# EPICS autosave request: iocs/motor/xps-ioc/db/XPSPositionCompare_settings.req
$(P)$(R)PositionCompareMode
$(P)$(R)PositionCompareMinPosition
$(P)$(R)PositionCompareMaxPosition
$(P)$(R)PositionCompareStepSize
$(P)$(R)PositionComparePulseWidth
$(P)$(R)PositionCompareSettlingTime
